(* IEC 61131-3 sources: repolevel_ST_code_completion/output/0122完整版本_无planner目前sota/repoeval_Proxy_Application/readful_result_before_fix, 2 files *)

(* ---- Proxy.st ---- *)
{attribute 'enable_dynamic_creation'}
FUNCTION_BLOCK Proxy IMPLEMENTS  Subject_Interface
VAR_INPUT
END_VAR
VAR_OUTPUT
END_VAR
VAR
    refToRealSubject : POINTER TO Realsubject;
    iTempPassword : INT;
END_VAR
VAR_STAT
    iRealPassword : INT := 1234;
END_VAR

METHOD fb_init
VAR_INPUT
    bInitRetains : BOOL;
    bInCopyCode : BOOL;
    ptrToRealSubject : POINTER TO Realsubject;
    iTempPassword : INT;
    iSetValue : INT;
    bReadWrite : BOOL;
END_VAR
VAR_OUTPUT
END_VAR
VAR
    refToRealSubject : POINTER TO Realsubject;
    iTempPassword : INT;
END_VAR
VAR_STAT
END_VAR

IF ptrToRealSubject <> 0 THEN
    refToRealSubject := ptrToRealSubject;
END_IF

IF bReadWrite THEN
    IF iTempPassword = iRealPassword THEN
        refToRealSubject^.iProp := iSetValue;
    END_IF
ELSE
    IF iTempPassword = iRealPassword THEN
        RETURN refToRealSubject^.iProp;
    ELSE
        RETURN -1; // Invalid password
    END_IF
END_IF
END_FUNCTION_BLOCK

(* ---- Realsubject.st ---- *)
{attribute 'enable_dynamic_creation'}
FUNCTION_BLOCK Realsubject IMPLEMENTS  Subject_Interface
VAR_INPUT
END_VAR
VAR_OUTPUT
END_VAR
VAR
    // Variable to get and set values
    iProp: INT;
END_VAR

VAR_STAT
END_VAR

METHOD PUBLIC Get_Method : INT
VAR
END_VAR
Get_Method := THIS^.iProp;

METHOD Set_Method
VAR_INPUT
    num : INT;
END_VAR
THIS^.iProp := num;
END_FUNCTION_BLOCK
